% RSLogix 500 project Robot Conveyor.RSS, saved by version 12.00.00.00 %
PROJECT "J14081"    % processor: MicroLogix 1400 %

PROGRAM FILES
  LAD 2   13 rungs
  LAD 3   7 rungs
  LAD 4   15 rungs
  LAD 5   12 rungs
  LAD 6   4 rungs
  LAD 7   6 rungs
  LAD 8   12 rungs

DATA FILES
  O0 OUTPUT  8 elements
  I1 INPUT  10 elements
  S2 STATUS  66 elements
  B3 BINARY  64 elements
  T4 TIMER  256 elements
  C5 COUNTER  1 elements
  R6 CONTROL  1 elements
  N7 INTEGER  1 elements
  F8 FLOAT  1 elements
  B9   16 elements
  B10   16 elements
  T11   32 elements
  T12   32 elements
  B13   16 elements
  B14   16 elements
  MG15   1 elements
  RI16   16 elements
  MG17   1 elements
  RI18   16 elements
  B33   16 elements

LADDER 2
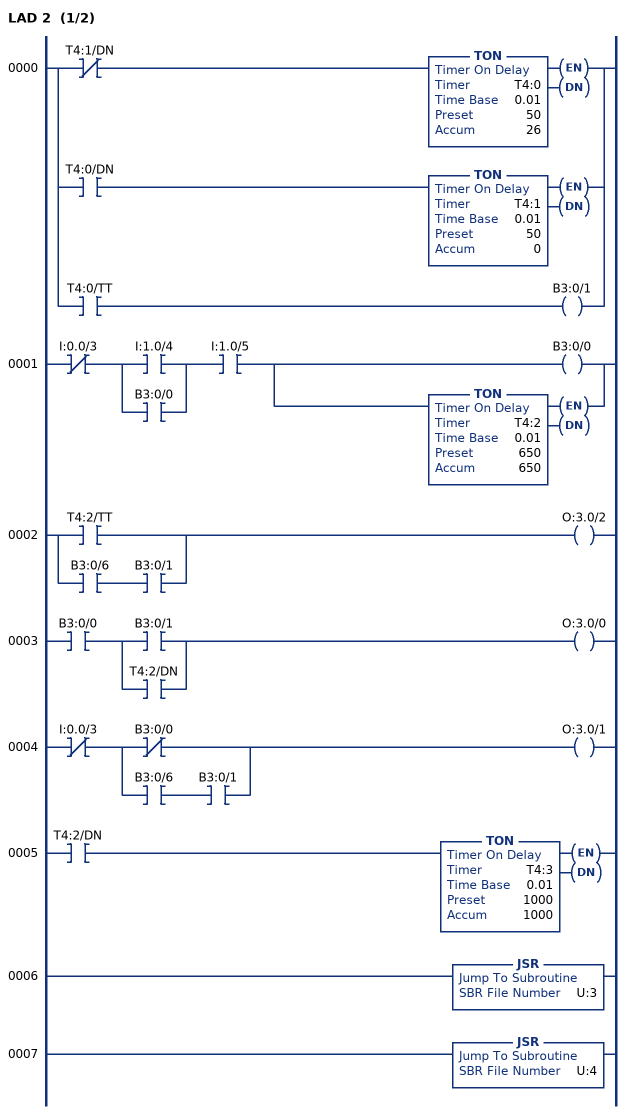
% Rung: 0 %
SOR BST XIO T4:1/DN TON T4:0 0.01 50 26 NXB XIC T4:0/DN TON T4:1 0.01 50 0 NXB XIC T4:0/TT OTE B3:0/1 BND EOR
% Rung: 1 %
SOR XIO I:0.0/3 BST XIC I:1.0/4 NXB XIC B3:0/0 BND XIC I:1.0/5 BST OTE B3:0/0 NXB TON T4:2 0.01 650 650 BND EOR
% Rung: 2 %
SOR BST XIC T4:2/TT NXB XIC B3:0/6 XIC B3:0/1 BND OTE O:3.0/2 EOR
% Rung: 3 %
SOR XIC B3:0/0 BST XIC B3:0/1 NXB XIC T4:2/DN BND OTE O:3.0/0 EOR
% Rung: 4 %
SOR XIO I:0.0/3 BST XIO B3:0/0 NXB XIC B3:0/6 XIC B3:0/1 BND OTE O:3.0/1 EOR
% Rung: 5 %
SOR XIC T4:2/DN TON T4:3 0.01 1000 1000 EOR
% Rung: 6 %
SOR JSR U:3 EOR
% Rung: 7 %
SOR JSR U:4 EOR

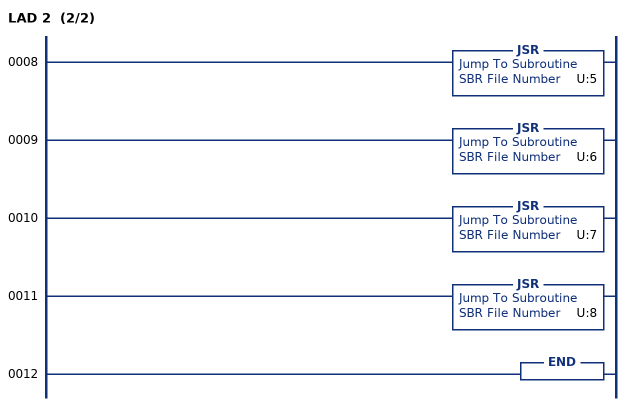
% Rung: 8 %
SOR JSR U:5 EOR
% Rung: 9 %
SOR JSR U:6 EOR
% Rung: 10 %
SOR JSR U:7 EOR
% Rung: 11 %
SOR JSR U:8 EOR
% Rung: 12 %
SOR END EOR

LADDER 3
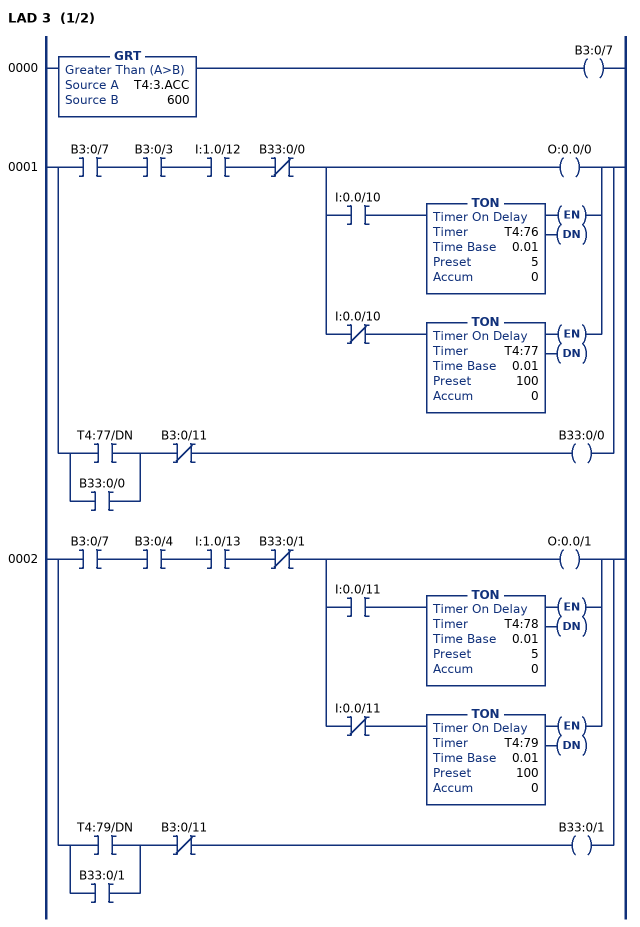
% Rung: 0 %
SOR GRT T4:3.ACC 600 OTE B3:0/7 EOR
% Rung: 1 %
SOR BST XIC B3:0/7 XIC B3:0/3 XIC I:1.0/12 XIO B33:0/0 BST OTE O:0.0/0 NXB XIC I:0.0/10 TON T4:76 0.01 5 0 NXB XIO I:0.0/10 TON T4:77 0.01 100 0 BND NXB BST XIC T4:77/DN NXB XIC B33:0/0 BND XIO B3:0/11 OTE B33:0/0 BND EOR
% Rung: 2 %
SOR BST XIC B3:0/7 XIC B3:0/4 XIC I:1.0/13 XIO B33:0/1 BST OTE O:0.0/1 NXB XIC I:0.0/11 TON T4:78 0.01 5 0 NXB XIO I:0.0/11 TON T4:79 0.01 100 0 BND NXB BST XIC T4:79/DN NXB XIC B33:0/1 BND XIO B3:0/11 OTE B33:0/1 BND EOR

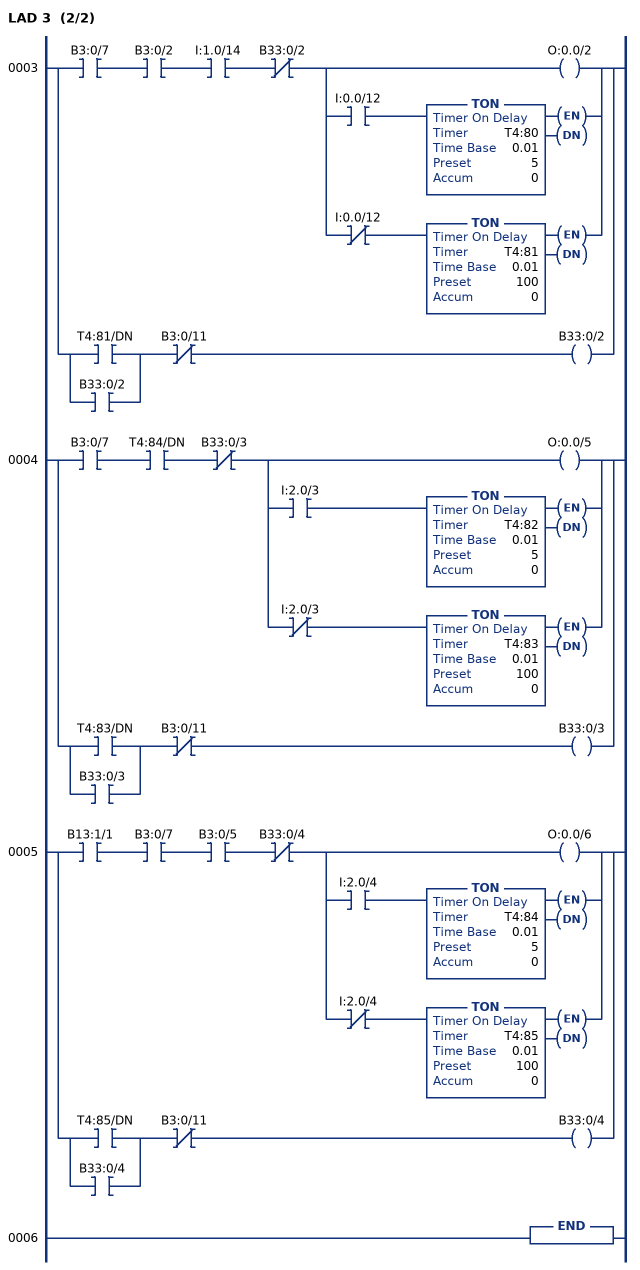
% Rung: 3 %
SOR BST XIC B3:0/7 XIC B3:0/2 XIC I:1.0/14 XIO B33:0/2 BST OTE O:0.0/2 NXB XIC I:0.0/12 TON T4:80 0.01 5 0 NXB XIO I:0.0/12 TON T4:81 0.01 100 0 BND NXB BST XIC T4:81/DN NXB XIC B33:0/2 BND XIO B3:0/11 OTE B33:0/2 BND EOR
% Rung: 4 %
SOR BST XIC B3:0/7 XIC T4:84/DN XIO B33:0/3 BST OTE O:0.0/5 NXB XIC I:2.0/3 TON T4:82 0.01 5 0 NXB XIO I:2.0/3 TON T4:83 0.01 100 0 BND NXB BST XIC T4:83/DN NXB XIC B33:0/3 BND XIO B3:0/11 OTE B33:0/3 BND EOR
% Rung: 5 %
SOR BST XIC B13:1/1 XIC B3:0/7 XIC B3:0/5 XIO B33:0/4 BST OTE O:0.0/6 NXB XIC I:2.0/4 TON T4:84 0.01 5 0 NXB XIO I:2.0/4 TON T4:85 0.01 100 0 BND NXB BST XIC T4:85/DN NXB XIC B33:0/4 BND XIO B3:0/11 OTE B33:0/4 BND EOR
% Rung: 6 %
SOR END EOR

LADDER 4
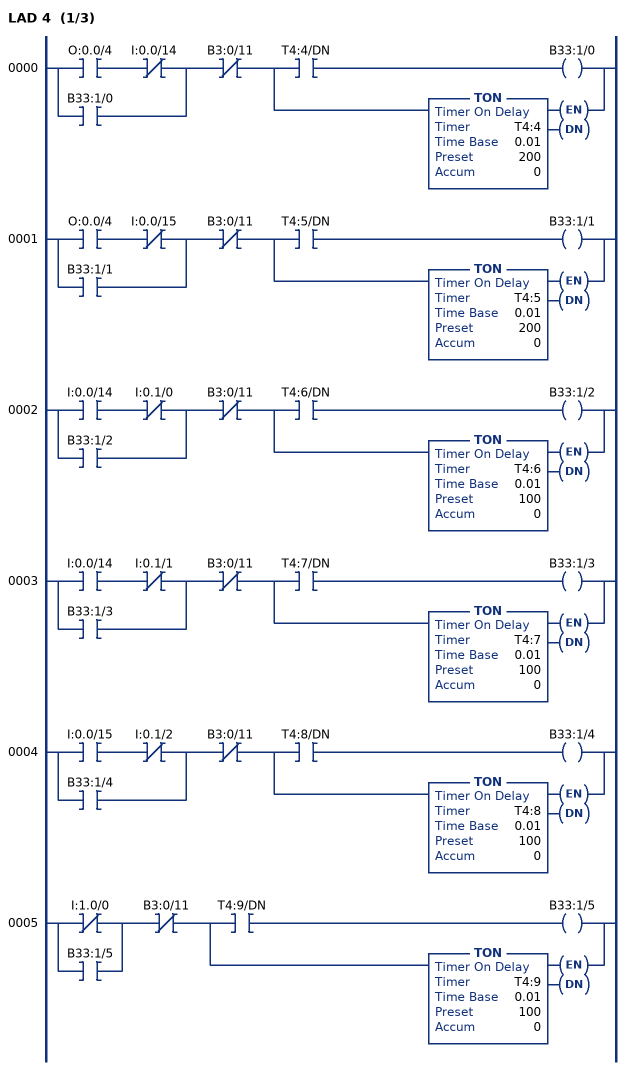
% Rung: 0 %
SOR BST XIC O:0.0/4 XIO I:0.0/14 NXB XIC B33:1/0 BND XIO B3:0/11 BST XIC T4:4/DN OTE B33:1/0 NXB TON T4:4 0.01 200 0 BND EOR
% Rung: 1 %
SOR BST XIC O:0.0/4 XIO I:0.0/15 NXB XIC B33:1/1 BND XIO B3:0/11 BST XIC T4:5/DN OTE B33:1/1 NXB TON T4:5 0.01 200 0 BND EOR
% Rung: 2 %
SOR BST XIC I:0.0/14 XIO I:0.1/0 NXB XIC B33:1/2 BND XIO B3:0/11 BST XIC T4:6/DN OTE B33:1/2 NXB TON T4:6 0.01 100 0 BND EOR
% Rung: 3 %
SOR BST XIC I:0.0/14 XIO I:0.1/1 NXB XIC B33:1/3 BND XIO B3:0/11 BST XIC T4:7/DN OTE B33:1/3 NXB TON T4:7 0.01 100 0 BND EOR
% Rung: 4 %
SOR BST XIC I:0.0/15 XIO I:0.1/2 NXB XIC B33:1/4 BND XIO B3:0/11 BST XIC T4:8/DN OTE B33:1/4 NXB TON T4:8 0.01 100 0 BND EOR
% Rung: 5 %
SOR BST XIO I:1.0/0 NXB XIC B33:1/5 BND XIO B3:0/11 BST XIC T4:9/DN OTE B33:1/5 NXB TON T4:9 0.01 100 0 BND EOR

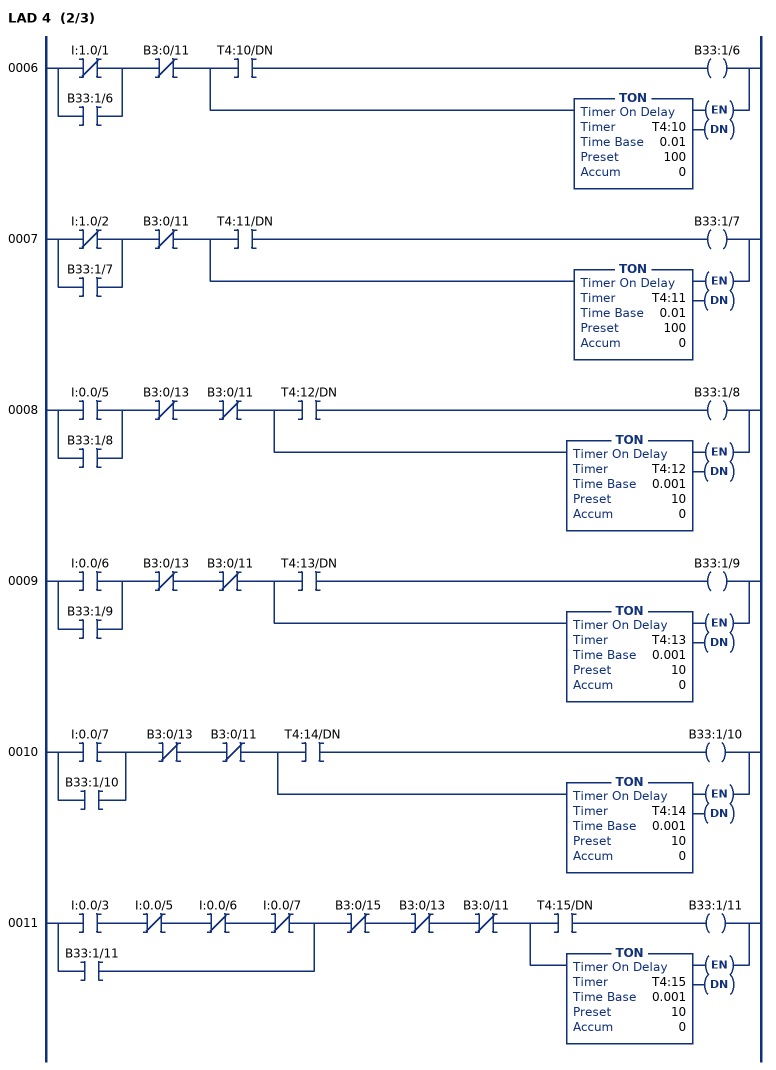
% Rung: 6 %
SOR BST XIO I:1.0/1 NXB XIC B33:1/6 BND XIO B3:0/11 BST XIC T4:10/DN OTE B33:1/6 NXB TON T4:10 0.01 100 0 BND EOR
% Rung: 7 %
SOR BST XIO I:1.0/2 NXB XIC B33:1/7 BND XIO B3:0/11 BST XIC T4:11/DN OTE B33:1/7 NXB TON T4:11 0.01 100 0 BND EOR
% Rung: 8 %
SOR BST XIC I:0.0/5 NXB XIC B33:1/8 BND XIO B3:0/13 XIO B3:0/11 BST XIC T4:12/DN OTE B33:1/8 NXB TON T4:12 0.001 10 0 BND EOR
% Rung: 9 %
SOR BST XIC I:0.0/6 NXB XIC B33:1/9 BND XIO B3:0/13 XIO B3:0/11 BST XIC T4:13/DN OTE B33:1/9 NXB TON T4:13 0.001 10 0 BND EOR
% Rung: 10 %
SOR BST XIC I:0.0/7 NXB XIC B33:1/10 BND XIO B3:0/13 XIO B3:0/11 BST XIC T4:14/DN OTE B33:1/10 NXB TON T4:14 0.001 10 0 BND EOR
% Rung: 11 %
SOR BST XIC I:0.0/3 XIO I:0.0/5 XIO I:0.0/6 XIO I:0.0/7 NXB XIC B33:1/11 BND XIO B3:0/15 XIO B3:0/13 XIO B3:0/11 BST XIC T4:15/DN OTE B33:1/11 NXB TON T4:15 0.001 10 0 BND EOR

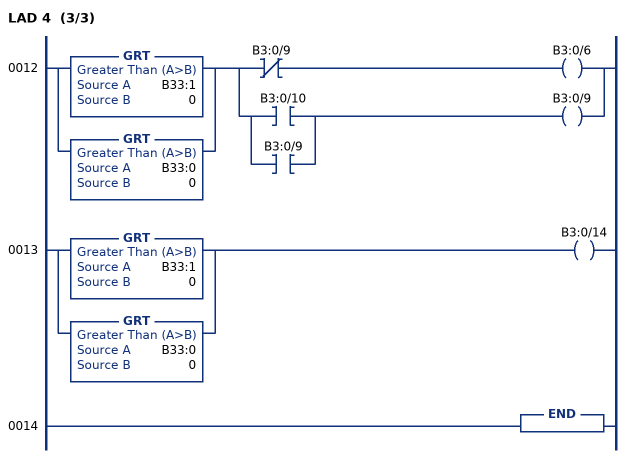
% Rung: 12 %
SOR BST GRT B33:1 0 NXB GRT B33:0 0 BND BST XIO B3:0/9 OTE B3:0/6 NXB BST XIC B3:0/10 NXB XIC B3:0/9 BND OTE B3:0/9 BND EOR
% Rung: 13 %
SOR BST GRT B33:1 0 NXB GRT B33:0 0 BND OTE B3:0/14 EOR
% Rung: 14 %
SOR END EOR

LADDER 5
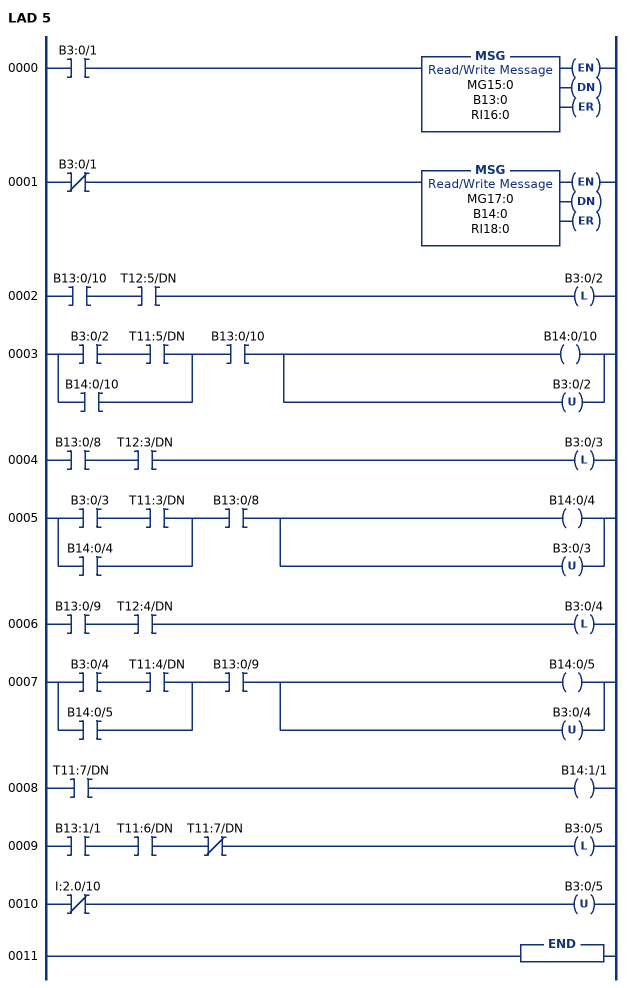
% Rung: 0 %
SOR XIC B3:0/1 MSG MG15:0 B13:0 RI16:0 EOR
%   MSG set-up: 500CPU Read | 33 | 16 | B13:0 | B13:0 | 0 | 0 | 0 | 192.168.1.101:0 | 0 | 0 | 192.168.1.101 | RI16:0 %
% Rung: 1 %
SOR XIO B3:0/1 MSG MG17:0 B14:0 RI18:0 EOR
%   MSG set-up: 500CPU Write | 33 | 16 | B14:0 | B14:0 | 0 | 0 | 0 | 192.168.1.101:0 | 0 | 0 | 192.168.1.101 | RI18:0 %
% Rung: 2 %
SOR XIC B13:0/10 XIC T12:5/DN OTL B3:0/2 EOR
% Rung: 3 %
SOR BST XIC B3:0/2 XIC T11:5/DN NXB XIC B14:0/10 BND XIC B13:0/10 BST OTE B14:0/10 NXB OTU B3:0/2 BND EOR
% Rung: 4 %
SOR XIC B13:0/8 XIC T12:3/DN OTL B3:0/3 EOR
% Rung: 5 %
SOR BST XIC B3:0/3 XIC T11:3/DN NXB XIC B14:0/4 BND XIC B13:0/8 BST OTE B14:0/4 NXB OTU B3:0/3 BND EOR
% Rung: 6 %
SOR XIC B13:0/9 XIC T12:4/DN OTL B3:0/4 EOR
% Rung: 7 %
SOR BST XIC B3:0/4 XIC T11:4/DN NXB XIC B14:0/5 BND XIC B13:0/9 BST OTE B14:0/5 NXB OTU B3:0/4 BND EOR
% Rung: 8 %
SOR XIC T11:7/DN OTE B14:1/1 EOR
% Rung: 9 %
SOR XIC B13:1/1 XIC T11:6/DN XIO T11:7/DN OTL B3:0/5 EOR
% Rung: 10 %
SOR XIO I:2.0/10 OTU B3:0/5 EOR
% Rung: 11 %
SOR END EOR

LADDER 6
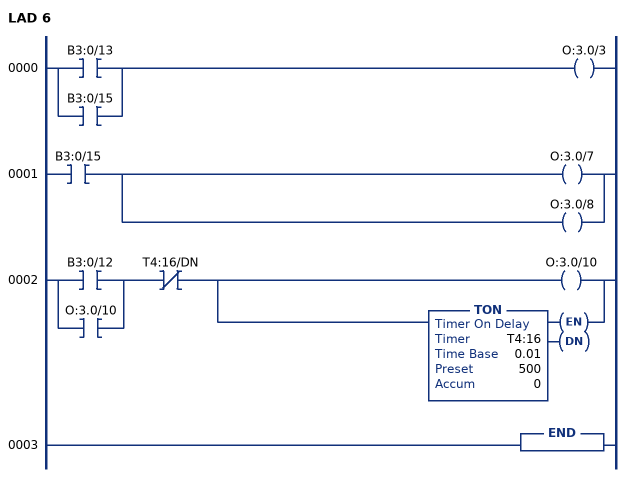
% Rung: 0 %
SOR BST XIC B3:0/13 NXB XIC B3:0/15 BND OTE O:3.0/3 EOR
% Rung: 1 %
SOR XIC B3:0/15 BST OTE O:3.0/7 NXB OTE O:3.0/8 BND EOR
% Rung: 2 %
SOR BST XIC B3:0/12 NXB XIC O:3.0/10 BND XIO T4:16/DN BST OTE O:3.0/10 NXB TON T4:16 0.01 500 0 BND EOR
% Rung: 3 %
SOR END EOR

LADDER 7
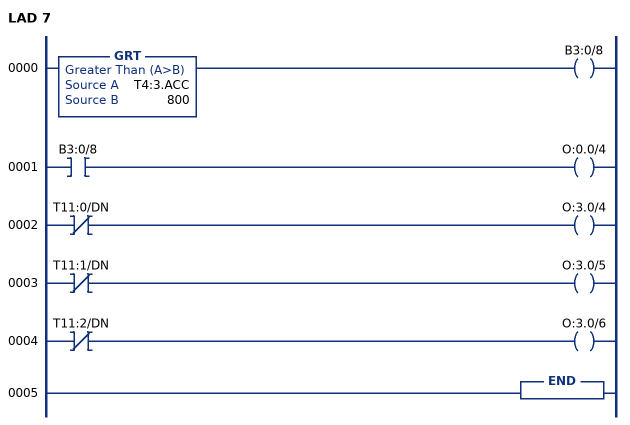
% Rung: 0 %
SOR GRT T4:3.ACC 800 OTE B3:0/8 EOR
% Rung: 1 %
SOR XIC B3:0/8 OTE O:0.0/4 EOR
% Rung: 2 %
SOR XIO T11:0/DN OTE O:3.0/4 EOR
% Rung: 3 %
SOR XIO T11:1/DN OTE O:3.0/5 EOR
% Rung: 4 %
SOR XIO T11:2/DN OTE O:3.0/6 EOR
% Rung: 5 %
SOR END EOR

LADDER 8
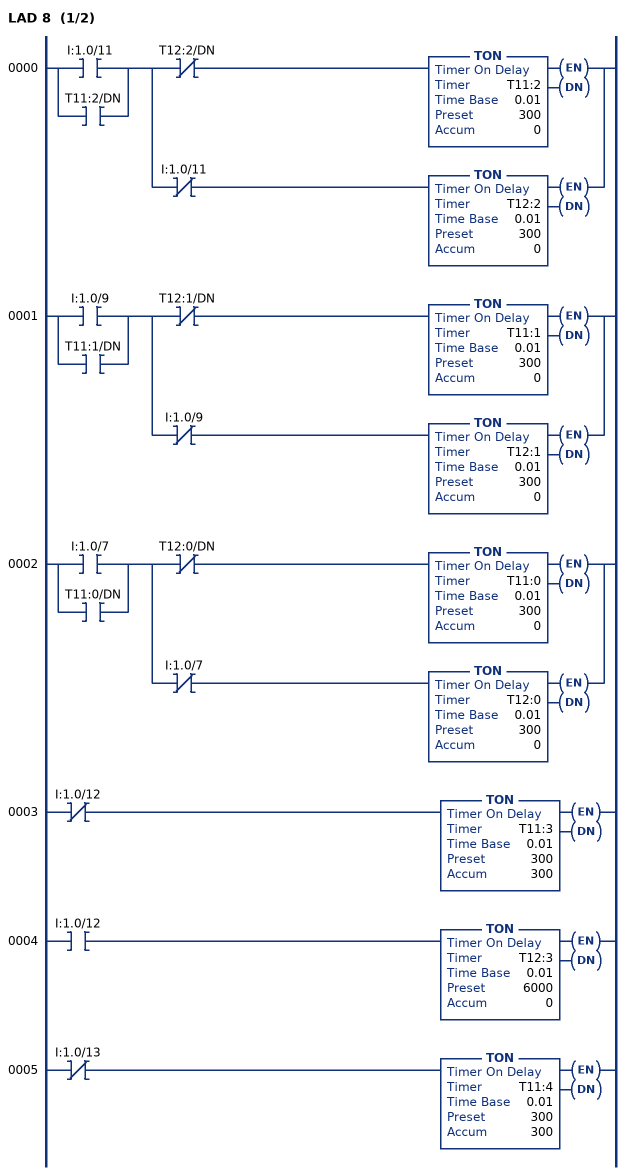
% Rung: 0 %
SOR BST XIC I:1.0/11 NXB XIC T11:2/DN BND BST XIO T12:2/DN TON T11:2 0.01 300 0 NXB XIO I:1.0/11 TON T12:2 0.01 300 0 BND EOR
% Rung: 1 %
SOR BST XIC I:1.0/9 NXB XIC T11:1/DN BND BST XIO T12:1/DN TON T11:1 0.01 300 0 NXB XIO I:1.0/9 TON T12:1 0.01 300 0 BND EOR
% Rung: 2 %
SOR BST XIC I:1.0/7 NXB XIC T11:0/DN BND BST XIO T12:0/DN TON T11:0 0.01 300 0 NXB XIO I:1.0/7 TON T12:0 0.01 300 0 BND EOR
% Rung: 3 %
SOR XIO I:1.0/12 TON T11:3 0.01 300 300 EOR
% Rung: 4 %
SOR XIC I:1.0/12 TON T12:3 0.01 6000 0 EOR
% Rung: 5 %
SOR XIO I:1.0/13 TON T11:4 0.01 300 300 EOR

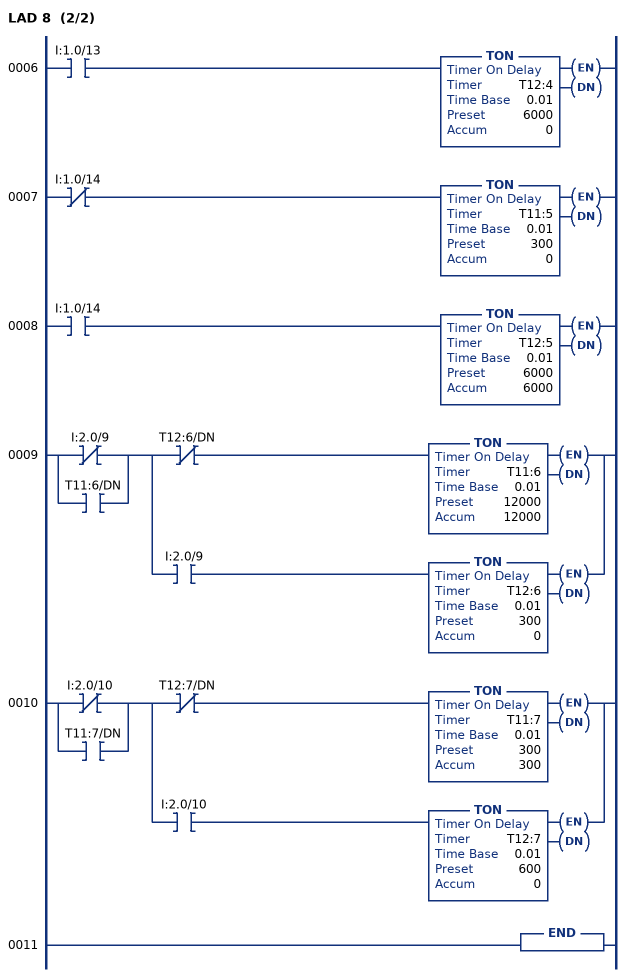
% Rung: 6 %
SOR XIC I:1.0/13 TON T12:4 0.01 6000 0 EOR
% Rung: 7 %
SOR XIO I:1.0/14 TON T11:5 0.01 300 0 EOR
% Rung: 8 %
SOR XIC I:1.0/14 TON T12:5 0.01 6000 6000 EOR
% Rung: 9 %
SOR BST XIO I:2.0/9 NXB XIC T11:6/DN BND BST XIO T12:6/DN TON T11:6 0.01 12000 12000 NXB XIC I:2.0/9 TON T12:6 0.01 300 0 BND EOR
% Rung: 10 %
SOR BST XIO I:2.0/10 NXB XIC T11:7/DN BND BST XIO T12:7/DN TON T11:7 0.01 300 300 NXB XIC I:2.0/10 TON T12:7 0.01 600 0 BND EOR
% Rung: 11 %
SOR END EOR

DATA TABLE (non-zero values as saved)
DATA B3
% B3:0 % 0X0183 0X0000 0X0000 0X0000 0X0000 0X0000 0X0000 0X0000 0X0000 0X0000
DATA T4
% .PRE .ACC %
% T4:0 % 50 26
% T4:1 % 50 0
% T4:2 % 650 650
% T4:3 % 1000 1000
% T4:4 % 200 0
% T4:5 % 200 0
% T4:6 % 100 0
% T4:7 % 100 0
% T4:8 % 100 0
% T4:9 % 100 0
% T4:10 % 100 0
% T4:11 % 100 0
% T4:12 % 10 0
% T4:13 % 10 0
% T4:14 % 10 0
% T4:15 % 10 0
% T4:16 % 500 0
% T4:76 % 5 0
% T4:77 % 100 0
% T4:78 % 5 0
% T4:79 % 100 0
% T4:80 % 5 0
% T4:81 % 100 0
% T4:82 % 5 0
% T4:83 % 100 0
% T4:84 % 5 0
% T4:85 % 100 0
DATA T11
% .PRE .ACC %
% T11:0 % 300 0
% T11:1 % 300 0
% T11:2 % 300 0
% T11:3 % 300 300
% T11:4 % 300 300
% T11:5 % 300 0
% T11:6 % 12000 12000
% T11:7 % 300 300
DATA T12
% .PRE .ACC %
% T12:0 % 300 0
% T12:1 % 300 0
% T12:2 % 300 0
% T12:3 % 6000 0
% T12:4 % 6000 0
% T12:5 % 6000 6000
% T12:6 % 300 0
% T12:7 % 600 0
DATA B13
% B13:0 % 0X0000 0X0002 0X0000 0X0000 0X0000 0X0000 0X0000 0X0000 0X0000 0X0000
DATA B14
% B14:0 % 0X0000 0X0002 0X0000 0X0000 0X0000 0X0000 0X0000 0X0000 0X0000 0X0000
